Yaskawa INFORM job: OVERLAP2.JBI

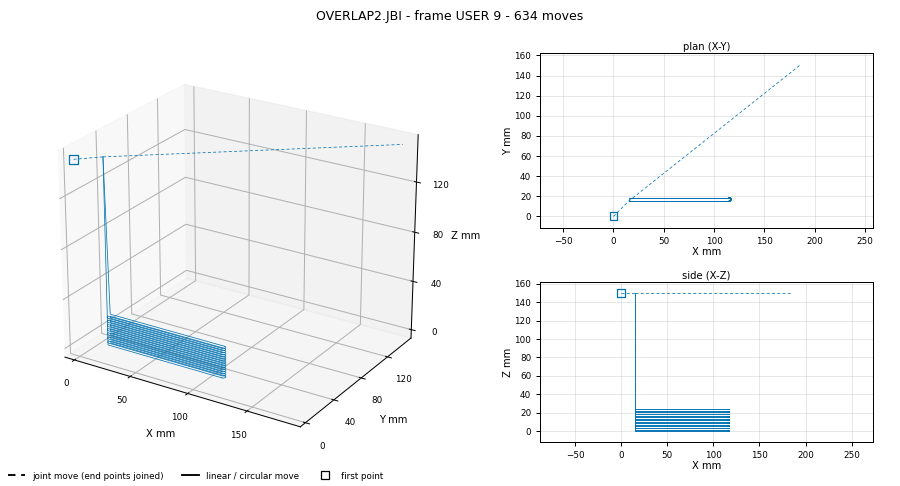
[picture p0: tool path of OVERLAP2.JBI in frame USER 9, 634 of 649 moves have a stored position in this frame; points joined in program order, loops and branches not executed]
/JOB
//NAME OVERLAP1
//POS
///NPOS 649,0,0,0,0,0
///USER 9
///TOOL 1
///POSTYPE USER
///RECTAN
///RCONF 1,0,0,0,0,0,0,0,0,0,0,0,0,0,0,0,0,0,0,0,0,0,0,0
C00000=0.000,0.000,150.000,0.0000,0.0000,-170.0000
C00001=15.000,15.000,150.000,0.0000,0.0000,-170.0000
C00002=15.000,15.000,0.000,0.0000,0.0000,-170.0000
C00003=20.000,15.000,0.000,0.0000,0.0000,-170.0000
C00004=25.000,15.000,0.000,0.0000,0.0000,-170.0000
C00005=30.000,15.000,0.000,0.0000,0.0000,-170.0000
C00006=35.000,15.000,0.000,0.0000,0.0000,-170.0000
C00007=40.000,15.000,0.000,0.0000,0.0000,-170.0000
C00008=45.000,15.000,0.000,0.0000,0.0000,-170.0000
C00009=50.000,15.000,0.000,0.0000,0.0000,-170.0000
C00010=55.000,15.000,0.000,0.0000,0.0000,-170.0000
C00011=60.000,15.000,0.000,0.0000,0.0000,-170.0000
C00012=65.000,15.000,0.000,0.0000,0.0000,-170.0000
C00013=70.000,15.000,0.000,0.0000,0.0000,-170.0000
C00014=75.000,15.000,0.000,0.0000,0.0000,-170.0000
C00015=80.000,15.000,0.000,0.0000,0.0000,-170.0000
C00016=85.000,15.000,0.000,0.0000,0.0000,-170.0000
C00017=90.000,15.000,0.000,0.0000,0.0000,-170.0000
C00018=95.000,15.000,0.000,0.0000,0.0000,-170.0000
C00019=100.000,15.000,0.000,0.0000,0.0000,-170.0000
C00020=105.000,15.000,0.000,0.0000,0.0000,-170.0000
C00021=110.000,15.000,0.000,0.0000,0.0000,-170.0000
C00022=115.000,15.000,0.000,0.0000,0.0000,-170.0000
C00023=116.875,16.875,0.000,0.0000,0.0000,-170.0000
C00024=115.000,18.750,0.000,0.0000,0.0000,-170.0000
C00025=110.000,18.750,0.000,0.0000,0.0000,-170.0000
C00026=105.000,18.750,0.000,0.0000,0.0000,-170.0000
C00027=100.000,18.750,0.000,0.0000,0.0000,-170.0000
C00028=95.000,18.750,0.000,0.0000,0.0000,-170.0000
C00029=90.000,18.750,0.000,0.0000,0.0000,-170.0000
C00030=85.000,18.750,0.000,0.0000,0.0000,-170.0000
C00031=80.000,18.750,0.000,0.0000,0.0000,-170.0000
C00032=75.000,18.750,0.000,0.0000,0.0000,-170.0000
C00033=70.000,18.750,0.000,0.0000,0.0000,-170.0000
C00034=65.000,18.750,0.000,0.0000,0.0000,-170.0000
C00035=60.000,18.750,0.000,0.0000,0.0000,-170.0000
C00036=55.000,18.750,0.000,0.0000,0.0000,-170.0000
C00037=50.000,18.750,0.000,0.0000,0.0000,-170.0000
C00038=45.000,18.750,0.000,0.0000,0.0000,-170.0000
C00039=40.000,18.750,0.000,0.0000,0.0000,-170.0000
C00040=35.000,18.750,0.000,0.0000,0.0000,-170.0000
C00041=30.000,18.750,0.000,0.0000,0.0000,-170.0000
C00042=25.000,18.750,0.000,0.0000,0.0000,-170.0000
C00043=20.000,18.750,0.000,0.0000,0.0000,-170.0000
C00044=15.000,18.750,0.000,0.0000,0.0000,-170.0000
C00045=15.000,18.750,1.700,0.0000,0.0000,-170.0000
C00046=20.000,18.750,1.700,0.0000,0.0000,-170.0000
C00047=25.000,18.750,1.700,0.0000,0.0000,-170.0000
C00048=30.000,18.750,1.700,0.0000,0.0000,-170.0000
C00049=35.000,18.750,1.700,0.0000,0.0000,-170.0000
C00050=40.000,18.750,1.700,0.0000,0.0000,-170.0000
C00051=45.000,18.750,1.700,0.0000,0.0000,-170.0000
C00052=50.000,18.750,1.700,0.0000,0.0000,-170.0000
C00053=55.000,18.750,1.700,0.0000,0.0000,-170.0000
C00054=60.000,18.750,1.700,0.0000,0.0000,-170.0000
C00055=65.000,18.750,1.700,0.0000,0.0000,-170.0000
C00056=70.000,18.750,1.700,0.0000,0.0000,-170.0000
C00057=75.000,18.750,1.700,0.0000,0.0000,-170.0000
C00058=80.000,18.750,1.700,0.0000,0.0000,-170.0000
C00059=85.000,18.750,1.700,0.0000,0.0000,-170.0000
C00060=90.000,18.750,1.700,0.0000,0.0000,-170.0000
C00061=95.000,18.750,1.700,0.0000,0.0000,-170.0000
C00062=100.000,18.750,1.700,0.0000,0.0000,-170.0000
C00063=105.000,18.750,1.700,0.0000,0.0000,-170.0000
C00064=110.000,18.750,1.700,0.0000,0.0000,-170.0000
C00065=115.000,18.750,1.700,0.0000,0.0000,-170.0000
C00066=116.875,16.875,1.700,0.0000,0.0000,-170.0000
C00067=115.000,15.000,1.700,0.0000,0.0000,-170.0000
C00068=110.000,15.000,1.700,0.0000,0.0000,-170.0000
C00069=105.000,15.000,1.700,0.0000,0.0000,-170.0000
C00070=100.000,15.000,1.700,0.0000,0.0000,-170.0000
C00071=95.000,15.000,1.700,0.0000,0.0000,-170.0000
C00072=90.000,15.000,1.700,0.0000,0.0000,-170.0000
C00073=85.000,15.000,1.700,0.0000,0.0000,-170.0000
C00074=80.000,15.000,1.700,0.0000,0.0000,-170.0000
C00075=75.000,15.000,1.700,0.0000,0.0000,-170.0000
C00076=70.000,15.000,1.700,0.0000,0.0000,-170.0000
C00077=65.000,15.000,1.700,0.0000,0.0000,-170.0000
C00078=60.000,15.000,1.700,0.0000,0.0000,-170.0000
C00079=55.000,15.000,1.700,0.0000,0.0000,-170.0000
C00080=50.000,15.000,1.700,0.0000,0.0000,-170.0000
C00081=45.000,15.000,1.700,0.0000,0.0000,-170.0000
C00082=40.000,15.000,1.700,0.0000,0.0000,-170.0000
C00083=35.000,15.000,1.700,0.0000,0.0000,-170.0000
C00084=30.000,15.000,1.700,0.0000,0.0000,-170.0000
C00085=25.000,15.000,1.700,0.0000,0.0000,-170.0000
C00086=20.000,15.000,1.700,0.0000,0.0000,-170.0000
C00087=15.000,15.000,1.700,0.0000,0.0000,-170.0000
C00088=15.000,15.000,3.400,0.0000,0.0000,-170.0000
C00089=20.000,15.000,3.400,0.0000,0.0000,-170.0000
C00090=25.000,15.000,3.400,0.0000,0.0000,-170.0000
C00091=30.000,15.000,3.400,0.0000,0.0000,-170.0000
C00092=35.000,15.000,3.400,0.0000,0.0000,-170.0000
C00093=40.000,15.000,3.400,0.0000,0.0000,-170.0000
C00094=45.000,15.000,3.400,0.0000,0.0000,-170.0000
C00095=50.000,15.000,3.400,0.0000,0.0000,-170.0000
C00096=55.000,15.000,3.400,0.0000,0.0000,-170.0000
C00097=60.000,15.000,3.400,0.0000,0.0000,-170.0000
C00098=65.000,15.000,3.400,0.0000,0.0000,-170.0000
C00099=70.000,15.000,3.400,0.0000,0.0000,-170.0000
C00100=75.000,15.000,3.400,0.0000,0.0000,-170.0000
C00101=80.000,15.000,3.400,0.0000,0.0000,-170.0000
C00102=85.000,15.000,3.400,0.0000,0.0000,-170.0000
C00103=90.000,15.000,3.400,0.0000,0.0000,-170.0000
C00104=95.000,15.000,3.400,0.0000,0.0000,-170.0000
C00105=100.000,15.000,3.400,0.0000,0.0000,-170.0000
C00106=105.000,15.000,3.400,0.0000,0.0000,-170.0000
C00107=110.000,15.000,3.400,0.0000,0.0000,-170.0000
C00108=115.000,15.000,3.400,0.0000,0.0000,-170.0000
C00109=116.875,16.875,3.400,0.0000,0.0000,-170.0000
C00110=115.000,18.750,3.400,0.0000,0.0000,-170.0000
C00111=110.000,18.750,3.400,0.0000,0.0000,-170.0000
C00112=105.000,18.750,3.400,0.0000,0.0000,-170.0000
C00113=100.000,18.750,3.400,0.0000,0.0000,-170.0000
C00114=95.000,18.750,3.400,0.0000,0.0000,-170.0000
C00115=90.000,18.750,3.400,0.0000,0.0000,-170.0000
C00116=85.000,18.750,3.400,0.0000,0.0000,-170.0000
C00117=80.000,18.750,3.400,0.0000,0.0000,-170.0000
C00118=75.000,18.750,3.400,0.0000,0.0000,-170.0000
C00119=70.000,18.750,3.400,0.0000,0.0000,-170.0000
C00120=65.000,18.750,3.400,0.0000,0.0000,-170.0000
C00121=60.000,18.750,3.400,0.0000,0.0000,-170.0000
C00122=55.000,18.750,3.400,0.0000,0.0000,-170.0000
C00123=50.000,18.750,3.400,0.0000,0.0000,-170.0000
C00124=45.000,18.750,3.400,0.0000,0.0000,-170.0000
C00125=40.000,18.750,3.400,0.0000,0.0000,-170.0000
C00126=35.000,18.750,3.400,0.0000,0.0000,-170.0000
C00127=30.000,18.750,3.400,0.0000,0.0000,-170.0000
C00128=25.000,18.750,3.400,0.0000,0.0000,-170.0000
C00129=20.000,18.750,3.400,0.0000,0.0000,-170.0000
C00130=15.000,18.750,3.400,0.0000,0.0000,-170.0000
C00131=15.000,18.750,5.100,0.0000,0.0000,-170.0000
C00132=20.000,18.750,5.100,0.0000,0.0000,-170.0000
C00133=25.000,18.750,5.100,0.0000,0.0000,-170.0000
C00134=30.000,18.750,5.100,0.0000,0.0000,-170.0000
C00135=35.000,18.750,5.100,0.0000,0.0000,-170.0000
C00136=40.000,18.750,5.100,0.0000,0.0000,-170.0000
C00137=45.000,18.750,5.100,0.0000,0.0000,-170.0000
C00138=50.000,18.750,5.100,0.0000,0.0000,-170.0000
C00139=55.000,18.750,5.100,0.0000,0.0000,-170.0000
C00140=60.000,18.750,5.100,0.0000,0.0000,-170.0000
C00141=65.000,18.750,5.100,0.0000,0.0000,-170.0000
C00142=70.000,18.750,5.100,0.0000,0.0000,-170.0000
C00143=75.000,18.750,5.100,0.0000,0.0000,-170.0000
C00144=80.000,18.750,5.100,0.0000,0.0000,-170.0000
C00145=85.000,18.750,5.100,0.0000,0.0000,-170.0000
C00146=90.000,18.750,5.100,0.0000,0.0000,-170.0000
C00147=95.000,18.750,5.100,0.0000,0.0000,-170.0000
C00148=100.000,18.750,5.100,0.0000,0.0000,-170.0000
C00149=105.000,18.750,5.100,0.0000,0.0000,-170.0000
C00150=110.000,18.750,5.100,0.0000,0.0000,-170.0000
C00151=115.000,18.750,5.100,0.0000,0.0000,-170.0000
C00152=116.875,16.875,5.100,0.0000,0.0000,-170.0000
C00153=115.000,15.000,5.100,0.0000,0.0000,-170.0000
C00154=110.000,15.000,5.100,0.0000,0.0000,-170.0000
C00155=105.000,15.000,5.100,0.0000,0.0000,-170.0000
C00156=100.000,15.000,5.100,0.0000,0.0000,-170.0000
C00157=95.000,15.000,5.100,0.0000,0.0000,-170.0000
C00158=90.000,15.000,5.100,0.0000,0.0000,-170.0000
C00159=85.000,15.000,5.100,0.0000,0.0000,-170.0000
C00160=80.000,15.000,5.100,0.0000,0.0000,-170.0000
C00161=75.000,15.000,5.100,0.0000,0.0000,-170.0000
C00162=70.000,15.000,5.100,0.0000,0.0000,-170.0000
C00163=65.000,15.000,5.100,0.0000,0.0000,-170.0000
C00164=60.000,15.000,5.100,0.0000,0.0000,-170.0000
C00165=55.000,15.000,5.100,0.0000,0.0000,-170.0000
C00166=50.000,15.000,5.100,0.0000,0.0000,-170.0000
C00167=45.000,15.000,5.100,0.0000,0.0000,-170.0000
C00168=40.000,15.000,5.100,0.0000,0.0000,-170.0000
C00169=35.000,15.000,5.100,0.0000,0.0000,-170.0000
C00170=30.000,15.000,5.100,0.0000,0.0000,-170.0000
C00171=25.000,15.000,5.100,0.0000,0.0000,-170.0000
C00172=20.000,15.000,5.100,0.0000,0.0000,-170.0000
C00173=15.000,15.000,5.100,0.0000,0.0000,-170.0000
C00174=15.000,15.000,6.800,0.0000,0.0000,-170.0000
C00175=20.000,15.000,6.800,0.0000,0.0000,-170.0000
C00176=25.000,15.000,6.800,0.0000,0.0000,-170.0000
C00177=30.000,15.000,6.800,0.0000,0.0000,-170.0000
C00178=35.000,15.000,6.800,0.0000,0.0000,-170.0000
C00179=40.000,15.000,6.800,0.0000,0.0000,-170.0000
C00180=45.000,15.000,6.800,0.0000,0.0000,-170.0000
C00181=50.000,15.000,6.800,0.0000,0.0000,-170.0000
C00182=55.000,15.000,6.800,0.0000,0.0000,-170.0000
C00183=60.000,15.000,6.800,0.0000,0.0000,-170.0000
C00184=65.000,15.000,6.800,0.0000,0.0000,-170.0000
C00185=70.000,15.000,6.800,0.0000,0.0000,-170.0000
C00186=75.000,15.000,6.800,0.0000,0.0000,-170.0000
C00187=80.000,15.000,6.800,0.0000,0.0000,-170.0000
C00188=85.000,15.000,6.800,0.0000,0.0000,-170.0000
C00189=90.000,15.000,6.800,0.0000,0.0000,-170.0000
C00190=95.000,15.000,6.800,0.0000,0.0000,-170.0000
C00191=100.000,15.000,6.800,0.0000,0.0000,-170.0000
C00192=105.000,15.000,6.800,0.0000,0.0000,-170.0000
C00193=110.000,15.000,6.800,0.0000,0.0000,-170.0000
C00194=115.000,15.000,6.800,0.0000,0.0000,-170.0000
C00195=116.875,16.875,6.800,0.0000,0.0000,-170.0000
C00196=115.000,18.750,6.800,0.0000,0.0000,-170.0000
C00197=110.000,18.750,6.800,0.0000,0.0000,-170.0000
C00198=105.000,18.750,6.800,0.0000,0.0000,-170.0000
C00199=100.000,18.750,6.800,0.0000,0.0000,-170.0000
C00200=95.000,18.750,6.800,0.0000,0.0000,-170.0000
C00201=90.000,18.750,6.800,0.0000,0.0000,-170.0000
C00202=85.000,18.750,6.800,0.0000,0.0000,-170.0000
C00203=80.000,18.750,6.800,0.0000,0.0000,-170.0000
C00204=75.000,18.750,6.800,0.0000,0.0000,-170.0000
C00205=70.000,18.750,6.800,0.0000,0.0000,-170.0000
C00206=65.000,18.750,6.800,0.0000,0.0000,-170.0000
C00207=60.000,18.750,6.800,0.0000,0.0000,-170.0000
C00208=55.000,18.750,6.800,0.0000,0.0000,-170.0000
C00209=50.000,18.750,6.800,0.0000,0.0000,-170.0000
C00210=45.000,18.750,6.800,0.0000,0.0000,-170.0000
C00211=40.000,18.750,6.800,0.0000,0.0000,-170.0000
C00212=35.000,18.750,6.800,0.0000,0.0000,-170.0000
C00213=30.000,18.750,6.800,0.0000,0.0000,-170.0000
C00214=25.000,18.750,6.800,0.0000,0.0000,-170.0000
C00215=20.000,18.750,6.800,0.0000,0.0000,-170.0000
C00216=15.000,18.750,6.800,0.0000,0.0000,-170.0000
C00217=15.000,18.750,8.500,0.0000,0.0000,-170.0000
C00218=20.000,18.750,8.500,0.0000,0.0000,-170.0000
C00219=25.000,18.750,8.500,0.0000,0.0000,-170.0000
C00220=30.000,18.750,8.500,0.0000,0.0000,-170.0000
C00221=35.000,18.750,8.500,0.0000,0.0000,-170.0000
C00222=40.000,18.750,8.500,0.0000,0.0000,-170.0000
C00223=45.000,18.750,8.500,0.0000,0.0000,-170.0000
C00224=50.000,18.750,8.500,0.0000,0.0000,-170.0000
C00225=55.000,18.750,8.500,0.0000,0.0000,-170.0000
C00226=60.000,18.750,8.500,0.0000,0.0000,-170.0000
C00227=65.000,18.750,8.500,0.0000,0.0000,-170.0000
C00228=70.000,18.750,8.500,0.0000,0.0000,-170.0000
C00229=75.000,18.750,8.500,0.0000,0.0000,-170.0000
C00230=80.000,18.750,8.500,0.0000,0.0000,-170.0000
C00231=85.000,18.750,8.500,0.0000,0.0000,-170.0000
C00232=90.000,18.750,8.500,0.0000,0.0000,-170.0000
C00233=95.000,18.750,8.500,0.0000,0.0000,-170.0000
C00234=100.000,18.750,8.500,0.0000,0.0000,-170.0000
C00235=105.000,18.750,8.500,0.0000,0.0000,-170.0000
C00236=110.000,18.750,8.500,0.0000,0.0000,-170.0000
C00237=115.000,18.750,8.500,0.0000,0.0000,-170.0000
C00238=116.875,16.875,8.500,0.0000,0.0000,-170.0000
C00239=115.000,15.000,8.500,0.0000,0.0000,-170.0000
C00240=110.000,15.000,8.500,0.0000,0.0000,-170.0000
C00241=105.000,15.000,8.500,0.0000,0.0000,-170.0000
C00242=100.000,15.000,8.500,0.0000,0.0000,-170.0000
C00243=95.000,15.000,8.500,0.0000,0.0000,-170.0000
C00244=90.000,15.000,8.500,0.0000,0.0000,-170.0000
C00245=85.000,15.000,8.500,0.0000,0.0000,-170.0000
C00246=80.000,15.000,8.500,0.0000,0.0000,-170.0000
C00247=75.000,15.000,8.500,0.0000,0.0000,-170.0000
C00248=70.000,15.000,8.500,0.0000,0.0000,-170.0000
C00249=65.000,15.000,8.500,0.0000,0.0000,-170.0000
C00250=60.000,15.000,8.500,0.0000,0.0000,-170.0000
C00251=55.000,15.000,8.500,0.0000,0.0000,-170.0000
C00252=50.000,15.000,8.500,0.0000,0.0000,-170.0000
C00253=45.000,15.000,8.500,0.0000,0.0000,-170.0000
C00254=40.000,15.000,8.500,0.0000,0.0000,-170.0000
C00255=35.000,15.000,8.500,0.0000,0.0000,-170.0000
C00256=30.000,15.000,8.500,0.0000,0.0000,-170.0000
C00257=25.000,15.000,8.500,0.0000,0.0000,-170.0000
C00258=20.000,15.000,8.500,0.0000,0.0000,-170.0000
C00259=15.000,15.000,8.500,0.0000,0.0000,-170.0000
C00260=15.000,15.000,10.200,0.0000,0.0000,-170.0000
C00261=20.000,15.000,10.200,0.0000,0.0000,-170.0000
C00262=25.000,15.000,10.200,0.0000,0.0000,-170.0000
C00263=30.000,15.000,10.200,0.0000,0.0000,-170.0000
C00264=35.000,15.000,10.200,0.0000,0.0000,-170.0000
C00265=40.000,15.000,10.200,0.0000,0.0000,-170.0000
C00266=45.000,15.000,10.200,0.0000,0.0000,-170.0000
C00267=50.000,15.000,10.200,0.0000,0.0000,-170.0000
C00268=55.000,15.000,10.200,0.0000,0.0000,-170.0000
C00269=60.000,15.000,10.200,0.0000,0.0000,-170.0000
C00270=65.000,15.000,10.200,0.0000,0.0000,-170.0000
C00271=70.000,15.000,10.200,0.0000,0.0000,-170.0000
C00272=75.000,15.000,10.200,0.0000,0.0000,-170.0000
C00273=80.000,15.000,10.200,0.0000,0.0000,-170.0000
C00274=85.000,15.000,10.200,0.0000,0.0000,-170.0000
C00275=90.000,15.000,10.200,0.0000,0.0000,-170.0000
C00276=95.000,15.000,10.200,0.0000,0.0000,-170.0000
C00277=100.000,15.000,10.200,0.0000,0.0000,-170.0000
C00278=105.000,15.000,10.200,0.0000,0.0000,-170.0000
C00279=110.000,15.000,10.200,0.0000,0.0000,-170.0000
C00280=115.000,15.000,10.200,0.0000,0.0000,-170.0000
C00281=116.875,16.875,10.200,0.0000,0.0000,-170.0000
C00282=115.000,18.750,10.200,0.0000,0.0000,-170.0000
C00283=110.000,18.750,10.200,0.0000,0.0000,-170.0000
C00284=105.000,18.750,10.200,0.0000,0.0000,-170.0000
C00285=100.000,18.750,10.200,0.0000,0.0000,-170.0000
C00286=95.000,18.750,10.200,0.0000,0.0000,-170.0000
C00287=90.000,18.750,10.200,0.0000,0.0000,-170.0000
C00288=85.000,18.750,10.200,0.0000,0.0000,-170.0000
C00289=80.000,18.750,10.200,0.0000,0.0000,-170.0000
C00290=75.000,18.750,10.200,0.0000,0.0000,-170.0000
C00291=70.000,18.750,10.200,0.0000,0.0000,-170.0000
C00292=65.000,18.750,10.200,0.0000,0.0000,-170.0000
C00293=60.000,18.750,10.200,0.0000,0.0000,-170.0000
C00294=55.000,18.750,10.200,0.0000,0.0000,-170.0000
C00295=50.000,18.750,10.200,0.0000,0.0000,-170.0000
C00296=45.000,18.750,10.200,0.0000,0.0000,-170.0000
C00297=40.000,18.750,10.200,0.0000,0.0000,-170.0000
C00298=35.000,18.750,10.200,0.0000,0.0000,-170.0000
C00299=30.000,18.750,10.200,0.0000,0.0000,-170.0000
C00300=25.000,18.750,10.200,0.0000,0.0000,-170.0000
C00301=20.000,18.750,10.200,0.0000,0.0000,-170.0000
C00302=15.000,18.750,10.200,0.0000,0.0000,-170.0000
C00303=15.000,18.750,11.900,0.0000,0.0000,-170.0000
C00304=20.000,18.750,11.900,0.0000,0.0000,-170.0000
C00305=25.000,18.750,11.900,0.0000,0.0000,-170.0000
C00306=30.000,18.750,11.900,0.0000,0.0000,-170.0000
C00307=35.000,18.750,11.900,0.0000,0.0000,-170.0000
C00308=40.000,18.750,11.900,0.0000,0.0000,-170.0000
C00309=45.000,18.750,11.900,0.0000,0.0000,-170.0000
C00310=50.000,18.750,11.900,0.0000,0.0000,-170.0000
C00311=55.000,18.750,11.900,0.0000,0.0000,-170.0000
C00312=60.000,18.750,11.900,0.0000,0.0000,-170.0000
C00313=65.000,18.750,11.900,0.0000,0.0000,-170.0000
C00314=70.000,18.750,11.900,0.0000,0.0000,-170.0000
C00315=75.000,18.750,11.900,0.0000,0.0000,-170.0000
C00316=80.000,18.750,11.900,0.0000,0.0000,-170.0000
C00317=85.000,18.750,11.900,0.0000,0.0000,-170.0000
C00318=90.000,18.750,11.900,0.0000,0.0000,-170.0000
C00319=95.000,18.750,11.900,0.0000,0.0000,-170.0000
C00320=100.000,18.750,11.900,0.0000,0.0000,-170.0000
C00321=105.000,18.750,11.900,0.0000,0.0000,-170.0000
C00322=110.000,18.750,11.900,0.0000,0.0000,-170.0000
C00323=115.000,18.750,11.900,0.0000,0.0000,-170.0000
C00324=116.875,16.875,11.900,0.0000,0.0000,-170.0000
C00325=115.000,15.000,11.900,0.0000,0.0000,-170.0000
C00326=110.000,15.000,11.900,0.0000,0.0000,-170.0000
C00327=105.000,15.000,11.900,0.0000,0.0000,-170.0000
C00328=100.000,15.000,11.900,0.0000,0.0000,-170.0000
C00329=95.000,15.000,11.900,0.0000,0.0000,-170.0000
C00330=90.000,15.000,11.900,0.0000,0.0000,-170.0000
C00331=85.000,15.000,11.900,0.0000,0.0000,-170.0000
C00332=80.000,15.000,11.900,0.0000,0.0000,-170.0000
C00333=75.000,15.000,11.900,0.0000,0.0000,-170.0000
C00334=70.000,15.000,11.900,0.0000,0.0000,-170.0000
C00335=65.000,15.000,11.900,0.0000,0.0000,-170.0000
C00336=60.000,15.000,11.900,0.0000,0.0000,-170.0000
C00337=55.000,15.000,11.900,0.0000,0.0000,-170.0000
C00338=50.000,15.000,11.900,0.0000,0.0000,-170.0000
C00339=45.000,15.000,11.900,0.0000,0.0000,-170.0000
C00340=40.000,15.000,11.900,0.0000,0.0000,-170.0000
C00341=35.000,15.000,11.900,0.0000,0.0000,-170.0000
C00342=30.000,15.000,11.900,0.0000,0.0000,-170.0000
C00343=25.000,15.000,11.900,0.0000,0.0000,-170.0000
C00344=20.000,15.000,11.900,0.0000,0.0000,-170.0000
C00345=15.000,15.000,11.900,0.0000,0.0000,-170.0000
C00346=15.000,15.000,13.600,0.0000,0.0000,-170.0000
C00347=20.000,15.000,13.600,0.0000,0.0000,-170.0000
C00348=25.000,15.000,13.600,0.0000,0.0000,-170.0000
C00349=30.000,15.000,13.600,0.0000,0.0000,-170.0000
C00350=35.000,15.000,13.600,0.0000,0.0000,-170.0000
C00351=40.000,15.000,13.600,0.0000,0.0000,-170.0000
C00352=45.000,15.000,13.600,0.0000,0.0000,-170.0000
C00353=50.000,15.000,13.600,0.0000,0.0000,-170.0000
C00354=55.000,15.000,13.600,0.0000,0.0000,-170.0000
C00355=60.000,15.000,13.600,0.0000,0.0000,-170.0000
C00356=65.000,15.000,13.600,0.0000,0.0000,-170.0000
C00357=70.000,15.000,13.600,0.0000,0.0000,-170.0000
C00358=75.000,15.000,13.600,0.0000,0.0000,-170.0000
C00359=80.000,15.000,13.600,0.0000,0.0000,-170.0000
C00360=85.000,15.000,13.600,0.0000,0.0000,-170.0000
C00361=90.000,15.000,13.600,0.0000,0.0000,-170.0000
C00362=95.000,15.000,13.600,0.0000,0.0000,-170.0000
C00363=100.000,15.000,13.600,0.0000,0.0000,-170.0000
C00364=105.000,15.000,13.600,0.0000,0.0000,-170.0000
C00365=110.000,15.000,13.600,0.0000,0.0000,-170.0000
C00366=115.000,15.000,13.600,0.0000,0.0000,-170.0000
C00367=116.875,16.875,13.600,0.0000,0.0000,-170.0000
C00368=115.000,18.750,13.600,0.0000,0.0000,-170.0000
C00369=110.000,18.750,13.600,0.0000,0.0000,-170.0000
C00370=105.000,18.750,13.600,0.0000,0.0000,-170.0000
C00371=100.000,18.750,13.600,0.0000,0.0000,-170.0000
C00372=95.000,18.750,13.600,0.0000,0.0000,-170.0000
C00373=90.000,18.750,13.600,0.0000,0.0000,-170.0000
C00374=85.000,18.750,13.600,0.0000,0.0000,-170.0000
C00375=80.000,18.750,13.600,0.0000,0.0000,-170.0000
C00376=75.000,18.750,13.600,0.0000,0.0000,-170.0000
C00377=70.000,18.750,13.600,0.0000,0.0000,-170.0000
C00378=65.000,18.750,13.600,0.0000,0.0000,-170.0000
C00379=60.000,18.750,13.600,0.0000,0.0000,-170.0000
C00380=55.000,18.750,13.600,0.0000,0.0000,-170.0000
C00381=50.000,18.750,13.600,0.0000,0.0000,-170.0000
C00382=45.000,18.750,13.600,0.0000,0.0000,-170.0000
C00383=40.000,18.750,13.600,0.0000,0.0000,-170.0000
C00384=35.000,18.750,13.600,0.0000,0.0000,-170.0000
C00385=30.000,18.750,13.600,0.0000,0.0000,-170.0000
C00386=25.000,18.750,13.600,0.0000,0.0000,-170.0000
C00387=20.000,18.750,13.600,0.0000,0.0000,-170.0000
C00388=15.000,18.750,13.600,0.0000,0.0000,-170.0000
C00389=15.000,18.750,15.300,0.0000,0.0000,-170.0000
C00390=20.000,18.750,15.300,0.0000,0.0000,-170.0000
C00391=25.000,18.750,15.300,0.0000,0.0000,-170.0000
C00392=30.000,18.750,15.300,0.0000,0.0000,-170.0000
C00393=35.000,18.750,15.300,0.0000,0.0000,-170.0000
C00394=40.000,18.750,15.300,0.0000,0.0000,-170.0000
C00395=45.000,18.750,15.300,0.0000,0.0000,-170.0000
C00396=50.000,18.750,15.300,0.0000,0.0000,-170.0000
C00397=55.000,18.750,15.300,0.0000,0.0000,-170.0000
C00398=60.000,18.750,15.300,0.0000,0.0000,-170.0000
C00399=65.000,18.750,15.300,0.0000,0.0000,-170.0000
C00400=70.000,18.750,15.300,0.0000,0.0000,-170.0000
C00401=75.000,18.750,15.300,0.0000,0.0000,-170.0000
C00402=80.000,18.750,15.300,0.0000,0.0000,-170.0000
C00403=85.000,18.750,15.300,0.0000,0.0000,-170.0000
C00404=90.000,18.750,15.300,0.0000,0.0000,-170.0000
C00405=95.000,18.750,15.300,0.0000,0.0000,-170.0000
C00406=100.000,18.750,15.300,0.0000,0.0000,-170.0000
C00407=105.000,18.750,15.300,0.0000,0.0000,-170.0000
C00408=110.000,18.750,15.300,0.0000,0.0000,-170.0000
C00409=115.000,18.750,15.300,0.0000,0.0000,-170.0000
C00410=116.875,16.875,15.300,0.0000,0.0000,-170.0000
C00411=115.000,15.000,15.300,0.0000,0.0000,-170.0000
C00412=110.000,15.000,15.300,0.0000,0.0000,-170.0000
C00413=105.000,15.000,15.300,0.0000,0.0000,-170.0000
C00414=100.000,15.000,15.300,0.0000,0.0000,-170.0000
C00415=95.000,15.000,15.300,0.0000,0.0000,-170.0000
C00416=90.000,15.000,15.300,0.0000,0.0000,-170.0000
C00417=85.000,15.000,15.300,0.0000,0.0000,-170.0000
C00418=80.000,15.000,15.300,0.0000,0.0000,-170.0000
C00419=75.000,15.000,15.300,0.0000,0.0000,-170.0000
C00420=70.000,15.000,15.300,0.0000,0.0000,-170.0000
C00421=65.000,15.000,15.300,0.0000,0.0000,-170.0000
C00422=60.000,15.000,15.300,0.0000,0.0000,-170.0000
C00423=55.000,15.000,15.300,0.0000,0.0000,-170.0000
C00424=50.000,15.000,15.300,0.0000,0.0000,-170.0000
C00425=45.000,15.000,15.300,0.0000,0.0000,-170.0000
C00426=40.000,15.000,15.300,0.0000,0.0000,-170.0000
C00427=35.000,15.000,15.300,0.0000,0.0000,-170.0000
C00428=30.000,15.000,15.300,0.0000,0.0000,-170.0000
C00429=25.000,15.000,15.300,0.0000,0.0000,-170.0000
C00430=20.000,15.000,15.300,0.0000,0.0000,-170.0000
C00431=15.000,15.000,15.300,0.0000,0.0000,-170.0000
C00432=15.000,15.000,17.000,0.0000,0.0000,-170.0000
C00433=20.000,15.000,17.000,0.0000,0.0000,-170.0000
C00434=25.000,15.000,17.000,0.0000,0.0000,-170.0000
C00435=30.000,15.000,17.000,0.0000,0.0000,-170.0000
C00436=35.000,15.000,17.000,0.0000,0.0000,-170.0000
C00437=40.000,15.000,17.000,0.0000,0.0000,-170.0000
C00438=45.000,15.000,17.000,0.0000,0.0000,-170.0000
C00439=50.000,15.000,17.000,0.0000,0.0000,-170.0000
C00440=55.000,15.000,17.000,0.0000,0.0000,-170.0000
C00441=60.000,15.000,17.000,0.0000,0.0000,-170.0000
C00442=65.000,15.000,17.000,0.0000,0.0000,-170.0000
C00443=70.000,15.000,17.000,0.0000,0.0000,-170.0000
C00444=75.000,15.000,17.000,0.0000,0.0000,-170.0000
C00445=80.000,15.000,17.000,0.0000,0.0000,-170.0000
C00446=85.000,15.000,17.000,0.0000,0.0000,-170.0000
C00447=90.000,15.000,17.000,0.0000,0.0000,-170.0000
C00448=95.000,15.000,17.000,0.0000,0.0000,-170.0000
C00449=100.000,15.000,17.000,0.0000,0.0000,-170.0000
C00450=105.000,15.000,17.000,0.0000,0.0000,-170.0000
C00451=110.000,15.000,17.000,0.0000,0.0000,-170.0000
C00452=115.000,15.000,17.000,0.0000,0.0000,-170.0000
C00453=116.875,16.875,17.000,0.0000,0.0000,-170.0000
C00454=115.000,18.750,17.000,0.0000,0.0000,-170.0000
C00455=110.000,18.750,17.000,0.0000,0.0000,-170.0000
C00456=105.000,18.750,17.000,0.0000,0.0000,-170.0000
C00457=100.000,18.750,17.000,0.0000,0.0000,-170.0000
C00458=95.000,18.750,17.000,0.0000,0.0000,-170.0000
C00459=90.000,18.750,17.000,0.0000,0.0000,-170.0000
C00460=85.000,18.750,17.000,0.0000,0.0000,-170.0000
C00461=80.000,18.750,17.000,0.0000,0.0000,-170.0000
C00462=75.000,18.750,17.000,0.0000,0.0000,-170.0000
C00463=70.000,18.750,17.000,0.0000,0.0000,-170.0000
C00464=65.000,18.750,17.000,0.0000,0.0000,-170.0000
C00465=60.000,18.750,17.000,0.0000,0.0000,-170.0000
C00466=55.000,18.750,17.000,0.0000,0.0000,-170.0000
C00467=50.000,18.750,17.000,0.0000,0.0000,-170.0000
C00468=45.000,18.750,17.000,0.0000,0.0000,-170.0000
C00469=40.000,18.750,17.000,0.0000,0.0000,-170.0000
C00470=35.000,18.750,17.000,0.0000,0.0000,-170.0000
C00471=30.000,18.750,17.000,0.0000,0.0000,-170.0000
C00472=25.000,18.750,17.000,0.0000,0.0000,-170.0000
C00473=20.000,18.750,17.000,0.0000,0.0000,-170.0000
C00474=15.000,18.750,17.000,0.0000,0.0000,-170.0000
C00475=15.000,18.750,18.700,0.0000,0.0000,-170.0000
C00476=20.000,18.750,18.700,0.0000,0.0000,-170.0000
C00477=25.000,18.750,18.700,0.0000,0.0000,-170.0000
C00478=30.000,18.750,18.700,0.0000,0.0000,-170.0000
C00479=35.000,18.750,18.700,0.0000,0.0000,-170.0000
C00480=40.000,18.750,18.700,0.0000,0.0000,-170.0000
C00481=45.000,18.750,18.700,0.0000,0.0000,-170.0000
C00482=50.000,18.750,18.700,0.0000,0.0000,-170.0000
C00483=55.000,18.750,18.700,0.0000,0.0000,-170.0000
C00484=60.000,18.750,18.700,0.0000,0.0000,-170.0000
C00485=65.000,18.750,18.700,0.0000,0.0000,-170.0000
C00486=70.000,18.750,18.700,0.0000,0.0000,-170.0000
C00487=75.000,18.750,18.700,0.0000,0.0000,-170.0000
C00488=80.000,18.750,18.700,0.0000,0.0000,-170.0000
C00489=85.000,18.750,18.700,0.0000,0.0000,-170.0000
C00490=90.000,18.750,18.700,0.0000,0.0000,-170.0000
C00491=95.000,18.750,18.700,0.0000,0.0000,-170.0000
C00492=100.000,18.750,18.700,0.0000,0.0000,-170.0000
C00493=105.000,18.750,18.700,0.0000,0.0000,-170.0000
C00494=110.000,18.750,18.700,0.0000,0.0000,-170.0000
C00495=115.000,18.750,18.700,0.0000,0.0000,-170.0000
C00496=116.875,16.875,18.700,0.0000,0.0000,-170.0000
C00497=115.000,15.000,18.700,0.0000,0.0000,-170.0000
C00498=110.000,15.000,18.700,0.0000,0.0000,-170.0000
C00499=105.000,15.000,18.700,0.0000,0.0000,-170.0000
C00500=100.000,15.000,18.700,0.0000,0.0000,-170.0000
C00501=95.000,15.000,18.700,0.0000,0.0000,-170.0000
C00502=90.000,15.000,18.700,0.0000,0.0000,-170.0000
C00503=85.000,15.000,18.700,0.0000,0.0000,-170.0000
C00504=80.000,15.000,18.700,0.0000,0.0000,-170.0000
C00505=75.000,15.000,18.700,0.0000,0.0000,-170.0000
C00506=70.000,15.000,18.700,0.0000,0.0000,-170.0000
C00507=65.000,15.000,18.700,0.0000,0.0000,-170.0000
C00508=60.000,15.000,18.700,0.0000,0.0000,-170.0000
C00509=55.000,15.000,18.700,0.0000,0.0000,-170.0000
C00510=50.000,15.000,18.700,0.0000,0.0000,-170.0000
C00511=45.000,15.000,18.700,0.0000,0.0000,-170.0000
C00512=40.000,15.000,18.700,0.0000,0.0000,-170.0000
C00513=35.000,15.000,18.700,0.0000,0.0000,-170.0000
C00514=30.000,15.000,18.700,0.0000,0.0000,-170.0000
C00515=25.000,15.000,18.700,0.0000,0.0000,-170.0000
C00516=20.000,15.000,18.700,0.0000,0.0000,-170.0000
C00517=15.000,15.000,18.700,0.0000,0.0000,-170.0000
C00518=15.000,15.000,20.400,0.0000,0.0000,-170.0000
C00519=20.000,15.000,20.400,0.0000,0.0000,-170.0000
C00520=25.000,15.000,20.400,0.0000,0.0000,-170.0000
C00521=30.000,15.000,20.400,0.0000,0.0000,-170.0000
C00522=35.000,15.000,20.400,0.0000,0.0000,-170.0000
C00523=40.000,15.000,20.400,0.0000,0.0000,-170.0000
C00524=45.000,15.000,20.400,0.0000,0.0000,-170.0000
C00525=50.000,15.000,20.400,0.0000,0.0000,-170.0000
C00526=55.000,15.000,20.400,0.0000,0.0000,-170.0000
C00527=60.000,15.000,20.400,0.0000,0.0000,-170.0000
C00528=65.000,15.000,20.400,0.0000,0.0000,-170.0000
C00529=70.000,15.000,20.400,0.0000,0.0000,-170.0000
C00530=75.000,15.000,20.400,0.0000,0.0000,-170.0000
C00531=80.000,15.000,20.400,0.0000,0.0000,-170.0000
C00532=85.000,15.000,20.400,0.0000,0.0000,-170.0000
C00533=90.000,15.000,20.400,0.0000,0.0000,-170.0000
C00534=95.000,15.000,20.400,0.0000,0.0000,-170.0000
C00535=100.000,15.000,20.400,0.0000,0.0000,-170.0000
C00536=105.000,15.000,20.400,0.0000,0.0000,-170.0000
C00537=110.000,15.000,20.400,0.0000,0.0000,-170.0000
C00538=115.000,15.000,20.400,0.0000,0.0000,-170.0000
C00539=116.875,16.875,20.400,0.0000,0.0000,-170.0000
C00540=115.000,18.750,20.400,0.0000,0.0000,-170.0000
C00541=110.000,18.750,20.400,0.0000,0.0000,-170.0000
C00542=105.000,18.750,20.400,0.0000,0.0000,-170.0000
C00543=100.000,18.750,20.400,0.0000,0.0000,-170.0000
C00544=95.000,18.750,20.400,0.0000,0.0000,-170.0000
C00545=90.000,18.750,20.400,0.0000,0.0000,-170.0000
C00546=85.000,18.750,20.400,0.0000,0.0000,-170.0000
C00547=80.000,18.750,20.400,0.0000,0.0000,-170.0000
C00548=75.000,18.750,20.400,0.0000,0.0000,-170.0000
C00549=70.000,18.750,20.400,0.0000,0.0000,-170.0000
C00550=65.000,18.750,20.400,0.0000,0.0000,-170.0000
C00551=60.000,18.750,20.400,0.0000,0.0000,-170.0000
C00552=55.000,18.750,20.400,0.0000,0.0000,-170.0000
C00553=50.000,18.750,20.400,0.0000,0.0000,-170.0000
C00554=45.000,18.750,20.400,0.0000,0.0000,-170.0000
C00555=40.000,18.750,20.400,0.0000,0.0000,-170.0000
C00556=35.000,18.750,20.400,0.0000,0.0000,-170.0000
C00557=30.000,18.750,20.400,0.0000,0.0000,-170.0000
C00558=25.000,18.750,20.400,0.0000,0.0000,-170.0000
C00559=20.000,18.750,20.400,0.0000,0.0000,-170.0000
C00560=15.000,18.750,20.400,0.0000,0.0000,-170.0000
C00561=15.000,18.750,22.100,0.0000,0.0000,-170.0000
C00562=20.000,18.750,22.100,0.0000,0.0000,-170.0000
C00563=25.000,18.750,22.100,0.0000,0.0000,-170.0000
C00564=30.000,18.750,22.100,0.0000,0.0000,-170.0000
C00565=35.000,18.750,22.100,0.0000,0.0000,-170.0000
C00566=40.000,18.750,22.100,0.0000,0.0000,-170.0000
C00567=45.000,18.750,22.100,0.0000,0.0000,-170.0000
C00568=50.000,18.750,22.100,0.0000,0.0000,-170.0000
C00569=55.000,18.750,22.100,0.0000,0.0000,-170.0000
C00570=60.000,18.750,22.100,0.0000,0.0000,-170.0000
C00571=65.000,18.750,22.100,0.0000,0.0000,-170.0000
C00572=70.000,18.750,22.100,0.0000,0.0000,-170.0000
C00573=75.000,18.750,22.100,0.0000,0.0000,-170.0000
C00574=80.000,18.750,22.100,0.0000,0.0000,-170.0000
C00575=85.000,18.750,22.100,0.0000,0.0000,-170.0000
C00576=90.000,18.750,22.100,0.0000,0.0000,-170.0000
C00577=95.000,18.750,22.100,0.0000,0.0000,-170.0000
C00578=100.000,18.750,22.100,0.0000,0.0000,-170.0000
C00579=105.000,18.750,22.100,0.0000,0.0000,-170.0000
C00580=110.000,18.750,22.100,0.0000,0.0000,-170.0000
C00581=115.000,18.750,22.100,0.0000,0.0000,-170.0000
C00582=116.875,16.875,22.100,0.0000,0.0000,-170.0000
C00583=115.000,15.000,22.100,0.0000,0.0000,-170.0000
C00584=110.000,15.000,22.100,0.0000,0.0000,-170.0000
C00585=105.000,15.000,22.100,0.0000,0.0000,-170.0000
C00586=100.000,15.000,22.100,0.0000,0.0000,-170.0000
C00587=95.000,15.000,22.100,0.0000,0.0000,-170.0000
C00588=90.000,15.000,22.100,0.0000,0.0000,-170.0000
C00589=85.000,15.000,22.100,0.0000,0.0000,-170.0000
C00590=80.000,15.000,22.100,0.0000,0.0000,-170.0000
C00591=75.000,15.000,22.100,0.0000,0.0000,-170.0000
C00592=70.000,15.000,22.100,0.0000,0.0000,-170.0000
C00593=65.000,15.000,22.100,0.0000,0.0000,-170.0000
C00594=60.000,15.000,22.100,0.0000,0.0000,-170.0000
C00595=55.000,15.000,22.100,0.0000,0.0000,-170.0000
C00596=50.000,15.000,22.100,0.0000,0.0000,-170.0000
C00597=45.000,15.000,22.100,0.0000,0.0000,-170.0000
C00598=40.000,15.000,22.100,0.0000,0.0000,-170.0000
C00599=35.000,15.000,22.100,0.0000,0.0000,-170.0000
C00600=30.000,15.000,22.100,0.0000,0.0000,-170.0000
C00601=25.000,15.000,22.100,0.0000,0.0000,-170.0000
C00602=20.000,15.000,22.100,0.0000,0.0000,-170.0000
C00603=15.000,15.000,22.100,0.0000,0.0000,-170.0000
C00604=15.000,15.000,23.800,0.0000,0.0000,-170.0000
C00605=20.000,15.000,23.800,0.0000,0.0000,-170.0000
C00606=25.000,15.000,23.800,0.0000,0.0000,-170.0000
C00607=30.000,15.000,23.800,0.0000,0.0000,-170.0000
C00608=35.000,15.000,23.800,0.0000,0.0000,-170.0000
C00609=40.000,15.000,23.800,0.0000,0.0000,-170.0000
C00610=45.000,15.000,23.800,0.0000,0.0000,-170.0000
C00611=50.000,15.000,23.800,0.0000,0.0000,-170.0000
C00612=55.000,15.000,23.800,0.0000,0.0000,-170.0000
C00613=60.000,15.000,23.800,0.0000,0.0000,-170.0000
C00614=65.000,15.000,23.800,0.0000,0.0000,-170.0000
C00615=70.000,15.000,23.800,0.0000,0.0000,-170.0000
C00616=75.000,15.000,23.800,0.0000,0.0000,-170.0000
C00617=80.000,15.000,23.800,0.0000,0.0000,-170.0000
C00618=85.000,15.000,23.800,0.0000,0.0000,-170.0000
C00619=90.000,15.000,23.800,0.0000,0.0000,-170.0000
C00620=95.000,15.000,23.800,0.0000,0.0000,-170.0000
C00621=100.000,15.000,23.800,0.0000,0.0000,-170.0000
C00622=105.000,15.000,23.800,0.0000,0.0000,-170.0000
C00623=110.000,15.000,23.800,0.0000,0.0000,-170.0000
C00624=115.000,15.000,23.800,0.0000,0.0000,-170.0000
C00625=116.875,16.875,23.800,0.0000,0.0000,-170.0000
C00626=115.000,18.750,23.800,0.0000,0.0000,-170.0000
C00627=110.000,18.750,23.800,0.0000,0.0000,-170.0000
C00628=105.000,18.750,23.800,0.0000,0.0000,-170.0000
C00629=100.000,18.750,23.800,0.0000,0.0000,-170.0000
C00630=95.000,18.750,23.800,0.0000,0.0000,-170.0000
C00631=90.000,18.750,23.800,0.0000,0.0000,-170.0000
C00632=85.000,18.750,23.800,0.0000,0.0000,-170.0000
C00633=80.000,18.750,23.800,0.0000,0.0000,-170.0000
C00634=75.000,18.750,23.800,0.0000,0.0000,-170.0000
C00635=70.000,18.750,23.800,0.0000,0.0000,-170.0000
C00636=65.000,18.750,23.800,0.0000,0.0000,-170.0000
C00637=60.000,18.750,23.800,0.0000,0.0000,-170.0000
C00638=55.000,18.750,23.800,0.0000,0.0000,-170.0000
C00639=50.000,18.750,23.800,0.0000,0.0000,-170.0000
C00640=45.000,18.750,23.800,0.0000,0.0000,-170.0000
C00641=40.000,18.750,23.800,0.0000,0.0000,-170.0000
C00642=35.000,18.750,23.800,0.0000,0.0000,-170.0000
C00643=30.000,18.750,23.800,0.0000,0.0000,-170.0000
C00644=25.000,18.750,23.800,0.0000,0.0000,-170.0000
C00645=20.000,18.750,23.800,0.0000,0.0000,-170.0000
C00646=15.000,18.750,23.800,0.0000,0.0000,-170.0000
C00647=15.000,15.000,150.000,0.0000,0.0000,-170.0000
C00648=185.000,150.000,150.000,0.0000,0.0000,-170.0000
//INST
///DATE 2026/11/06 13:28
///ATTR SC,RW,RJ
////FRAME USER 9
///GROUP1 RB1
NOP
MOVJ C00000 VJ=0.78
MOVJ C00001 VJ=0.78
MOVL C00002 V=11.0 PL=0
*LAG1
MACRO1 MJ#(0) ARGF1
ARCON
MOVL C00003 V=7.0 PL=0
MOVL C00004 V=7.0 PL=0
MOVL C00005 V=7.0 PL=0
MOVL C00006 V=7.0 PL=0
MOVL C00007 V=7.0 PL=0
MOVL C00008 V=7.0 PL=0
MOVL C00009 V=7.0 PL=0
MOVL C00010 V=7.0 PL=0
MOVL C00011 V=7.0 PL=0
MOVL C00012 V=7.0 PL=0
MOVL C00013 V=7.0 PL=0
MOVL C00014 V=7.0 PL=0
MOVL C00015 V=7.0 PL=0
MOVL C00016 V=7.0 PL=0
MOVL C00017 V=7.0 PL=0
MOVL C00018 V=7.0 PL=0
MOVL C00019 V=7.0 PL=0
MOVL C00020 V=7.0 PL=0
MOVL C00021 V=7.0 PL=0
MOVC C00022 V=7.0 ACC=20 DEC=20
MOVC C00023 V=7.0 ACC=20 DEC=20
MOVC C00024 V=7.0 ACC=20 DEC=20
MOVL C00025 V=7.0 PL=0
MOVL C00026 V=7.0 PL=0
MOVL C00027 V=7.0 PL=0
MOVL C00028 V=7.0 PL=0
MOVL C00029 V=7.0 PL=0
MOVL C00030 V=7.0 PL=0
MOVL C00031 V=7.0 PL=0
MOVL C00032 V=7.0 PL=0
MOVL C00033 V=7.0 PL=0
MOVL C00034 V=7.0 PL=0
MOVL C00035 V=7.0 PL=0
MOVL C00036 V=7.0 PL=0
MOVL C00037 V=7.0 PL=0
MOVL C00038 V=7.0 PL=0
MOVL C00039 V=7.0 PL=0
MOVL C00040 V=7.0 PL=0
MOVL C00041 V=7.0 PL=0
MOVL C00042 V=7.0 PL=0
MOVL C00043 V=7.0 PL=0
MOVL C00044 V=7.0 PL=0
ARCOF
TIMER T=30.00
*LAG2
MOVL C00045 V=11.0 PL=0
MACRO1 MJ#(0) ARGF2
ARCON
MOVL C00046 V=7.0 PL=0
MOVL C00047 V=7.0 PL=0
MOVL C00048 V=7.0 PL=0
MOVL C00049 V=7.0 PL=0
MOVL C00050 V=7.0 PL=0
MOVL C00051 V=7.0 PL=0
MOVL C00052 V=7.0 PL=0
MOVL C00053 V=7.0 PL=0
MOVL C00054 V=7.0 PL=0
MOVL C00055 V=7.0 PL=0
MOVL C00056 V=7.0 PL=0
MOVL C00057 V=7.0 PL=0
MOVL C00058 V=7.0 PL=0
MOVL C00059 V=7.0 PL=0
MOVL C00060 V=7.0 PL=0
MOVL C00061 V=7.0 PL=0
MOVL C00062 V=7.0 PL=0
MOVL C00063 V=7.0 PL=0
MOVL C00064 V=7.0 PL=0
MOVC C00065 V=7.0 ACC=20 DEC=20
MOVC C00066 V=7.0 ACC=20 DEC=20
MOVC C00067 V=7.0 ACC=20 DEC=20
MOVL C00068 V=7.0 PL=0
MOVL C00069 V=7.0 PL=0
MOVL C00070 V=7.0 PL=0
MOVL C00071 V=7.0 PL=0
MOVL C00072 V=7.0 PL=0
MOVL C00073 V=7.0 PL=0
MOVL C00074 V=7.0 PL=0
MOVL C00075 V=7.0 PL=0
MOVL C00076 V=7.0 PL=0
MOVL C00077 V=7.0 PL=0
MOVL C00078 V=7.0 PL=0
MOVL C00079 V=7.0 PL=0
MOVL C00080 V=7.0 PL=0
MOVL C00081 V=7.0 PL=0
MOVL C00082 V=7.0 PL=0
MOVL C00083 V=7.0 PL=0
MOVL C00084 V=7.0 PL=0
MOVL C00085 V=7.0 PL=0
MOVL C00086 V=7.0 PL=0
MOVL C00087 V=7.0 PL=0
ARCOF
TIMER T=30.00
*LAG3
MOVL C00088 V=11.0 PL=0
MACRO1 MJ#(0) ARGF2
ARCON
MOVL C00089 V=7.0 PL=0
MOVL C00090 V=7.0 PL=0
MOVL C00091 V=7.0 PL=0
MOVL C00092 V=7.0 PL=0
MOVL C00093 V=7.0 PL=0
MOVL C00094 V=7.0 PL=0
MOVL C00095 V=7.0 PL=0
MOVL C00096 V=7.0 PL=0
MOVL C00097 V=7.0 PL=0
MOVL C00098 V=7.0 PL=0
MOVL C00099 V=7.0 PL=0
MOVL C00100 V=7.0 PL=0
MOVL C00101 V=7.0 PL=0
MOVL C00102 V=7.0 PL=0
MOVL C00103 V=7.0 PL=0
MOVL C00104 V=7.0 PL=0
MOVL C00105 V=7.0 PL=0
MOVL C00106 V=7.0 PL=0
MOVL C00107 V=7.0 PL=0
MOVC C00108 V=7.0 ACC=20 DEC=20
MOVC C00109 V=7.0 ACC=20 DEC=20
MOVC C00110 V=7.0 ACC=20 DEC=20
MOVL C00111 V=7.0 PL=0
MOVL C00112 V=7.0 PL=0
MOVL C00113 V=7.0 PL=0
MOVL C00114 V=7.0 PL=0
MOVL C00115 V=7.0 PL=0
MOVL C00116 V=7.0 PL=0
MOVL C00117 V=7.0 PL=0
MOVL C00118 V=7.0 PL=0
MOVL C00119 V=7.0 PL=0
MOVL C00120 V=7.0 PL=0
MOVL C00121 V=7.0 PL=0
MOVL C00122 V=7.0 PL=0
MOVL C00123 V=7.0 PL=0
MOVL C00124 V=7.0 PL=0
MOVL C00125 V=7.0 PL=0
MOVL C00126 V=7.0 PL=0
MOVL C00127 V=7.0 PL=0
MOVL C00128 V=7.0 PL=0
MOVL C00129 V=7.0 PL=0
MOVL C00130 V=7.0 PL=0
ARCOF
TIMER T=30.00
*LAG4
MOVL C00131 V=11.0 PL=0
MACRO1 MJ#(0) ARGF2
ARCON
MOVL C00132 V=7.0 PL=0
MOVL C00133 V=7.0 PL=0
MOVL C00134 V=7.0 PL=0
MOVL C00135 V=7.0 PL=0
MOVL C00136 V=7.0 PL=0
MOVL C00137 V=7.0 PL=0
MOVL C00138 V=7.0 PL=0
MOVL C00139 V=7.0 PL=0
MOVL C00140 V=7.0 PL=0
MOVL C00141 V=7.0 PL=0
MOVL C00142 V=7.0 PL=0
MOVL C00143 V=7.0 PL=0
MOVL C00144 V=7.0 PL=0
MOVL C00145 V=7.0 PL=0
MOVL C00146 V=7.0 PL=0
MOVL C00147 V=7.0 PL=0
MOVL C00148 V=7.0 PL=0
MOVL C00149 V=7.0 PL=0
MOVL C00150 V=7.0 PL=0
MOVC C00151 V=7.0 ACC=20 DEC=20
MOVC C00152 V=7.0 ACC=20 DEC=20
MOVC C00153 V=7.0 ACC=20 DEC=20
MOVL C00154 V=7.0 PL=0
MOVL C00155 V=7.0 PL=0
MOVL C00156 V=7.0 PL=0
MOVL C00157 V=7.0 PL=0
MOVL C00158 V=7.0 PL=0
MOVL C00159 V=7.0 PL=0
MOVL C00160 V=7.0 PL=0
MOVL C00161 V=7.0 PL=0
MOVL C00162 V=7.0 PL=0
MOVL C00163 V=7.0 PL=0
MOVL C00164 V=7.0 PL=0
MOVL C00165 V=7.0 PL=0
MOVL C00166 V=7.0 PL=0
MOVL C00167 V=7.0 PL=0
MOVL C00168 V=7.0 PL=0
MOVL C00169 V=7.0 PL=0
MOVL C00170 V=7.0 PL=0
MOVL C00171 V=7.0 PL=0
MOVL C00172 V=7.0 PL=0
MOVL C00173 V=7.0 PL=0
ARCOF
TIMER T=30.00
*LAG5
MOVL C00174 V=11.0 PL=0
MACRO1 MJ#(0) ARGF2
ARCON
MOVL C00175 V=7.0 PL=0
MOVL C00176 V=7.0 PL=0
MOVL C00177 V=7.0 PL=0
MOVL C00178 V=7.0 PL=0
MOVL C00179 V=7.0 PL=0
MOVL C00180 V=7.0 PL=0
MOVL C00181 V=7.0 PL=0
MOVL C00182 V=7.0 PL=0
MOVL C00183 V=7.0 PL=0
MOVL C00184 V=7.0 PL=0
MOVL C00185 V=7.0 PL=0
MOVL C00186 V=7.0 PL=0
MOVL C00187 V=7.0 PL=0
MOVL C00188 V=7.0 PL=0
MOVL C00189 V=7.0 PL=0
MOVL C00190 V=7.0 PL=0
MOVL C00191 V=7.0 PL=0
MOVL C00192 V=7.0 PL=0
MOVL C00193 V=7.0 PL=0
MOVC C00194 V=7.0 ACC=20 DEC=20
MOVC C00195 V=7.0 ACC=20 DEC=20
MOVC C00196 V=7.0 ACC=20 DEC=20
MOVL C00197 V=7.0 PL=0
MOVL C00198 V=7.0 PL=0
MOVL C00199 V=7.0 PL=0
MOVL C00200 V=7.0 PL=0
MOVL C00201 V=7.0 PL=0
MOVL C00202 V=7.0 PL=0
MOVL C00203 V=7.0 PL=0
MOVL C00204 V=7.0 PL=0
MOVL C00205 V=7.0 PL=0
MOVL C00206 V=7.0 PL=0
MOVL C00207 V=7.0 PL=0
MOVL C00208 V=7.0 PL=0
MOVL C00209 V=7.0 PL=0
MOVL C00210 V=7.0 PL=0
MOVL C00211 V=7.0 PL=0
MOVL C00212 V=7.0 PL=0
MOVL C00213 V=7.0 PL=0
MOVL C00214 V=7.0 PL=0
MOVL C00215 V=7.0 PL=0
MOVL C00216 V=7.0 PL=0
ARCOF
TIMER T=30.00
*LAG6
MOVL C00217 V=11.0 PL=0
MACRO1 MJ#(0) ARGF2
ARCON
MOVL C00218 V=7.0 PL=0
MOVL C00219 V=7.0 PL=0
MOVL C00220 V=7.0 PL=0
MOVL C00221 V=7.0 PL=0
MOVL C00222 V=7.0 PL=0
MOVL C00223 V=7.0 PL=0
MOVL C00224 V=7.0 PL=0
MOVL C00225 V=7.0 PL=0
MOVL C00226 V=7.0 PL=0
MOVL C00227 V=7.0 PL=0
MOVL C00228 V=7.0 PL=0
MOVL C00229 V=7.0 PL=0
MOVL C00230 V=7.0 PL=0
MOVL C00231 V=7.0 PL=0
MOVL C00232 V=7.0 PL=0
MOVL C00233 V=7.0 PL=0
MOVL C00234 V=7.0 PL=0
MOVL C00235 V=7.0 PL=0
MOVL C00236 V=7.0 PL=0
MOVC C00237 V=7.0 ACC=20 DEC=20
MOVC C00238 V=7.0 ACC=20 DEC=20
MOVC C00239 V=7.0 ACC=20 DEC=20
MOVL C00240 V=7.0 PL=0
MOVL C00241 V=7.0 PL=0
MOVL C00242 V=7.0 PL=0
MOVL C00243 V=7.0 PL=0
MOVL C00244 V=7.0 PL=0
MOVL C00245 V=7.0 PL=0
MOVL C00246 V=7.0 PL=0
MOVL C00247 V=7.0 PL=0
MOVL C00248 V=7.0 PL=0
MOVL C00249 V=7.0 PL=0
MOVL C00250 V=7.0 PL=0
MOVL C00251 V=7.0 PL=0
MOVL C00252 V=7.0 PL=0
MOVL C00253 V=7.0 PL=0
MOVL C00254 V=7.0 PL=0
MOVL C00255 V=7.0 PL=0
MOVL C00256 V=7.0 PL=0
MOVL C00257 V=7.0 PL=0
MOVL C00258 V=7.0 PL=0
MOVL C00259 V=7.0 PL=0
ARCOF
TIMER T=30.00
*LAG7
MOVL C00260 V=11.0 PL=0
MACRO1 MJ#(0) ARGF2
ARCON
MOVL C00261 V=7.0 PL=0
MOVL C00262 V=7.0 PL=0
MOVL C00263 V=7.0 PL=0
MOVL C00264 V=7.0 PL=0
MOVL C00265 V=7.0 PL=0
MOVL C00266 V=7.0 PL=0
MOVL C00267 V=7.0 PL=0
MOVL C00268 V=7.0 PL=0
MOVL C00269 V=7.0 PL=0
MOVL C00270 V=7.0 PL=0
MOVL C00271 V=7.0 PL=0
MOVL C00272 V=7.0 PL=0
MOVL C00273 V=7.0 PL=0
MOVL C00274 V=7.0 PL=0
MOVL C00275 V=7.0 PL=0
MOVL C00276 V=7.0 PL=0
MOVL C00277 V=7.0 PL=0
MOVL C00278 V=7.0 PL=0
MOVL C00279 V=7.0 PL=0
MOVC C00280 V=7.0 ACC=20 DEC=20
MOVC C00281 V=7.0 ACC=20 DEC=20
MOVC C00282 V=7.0 ACC=20 DEC=20
MOVL C00283 V=7.0 PL=0
MOVL C00284 V=7.0 PL=0
MOVL C00285 V=7.0 PL=0
MOVL C00286 V=7.0 PL=0
MOVL C00287 V=7.0 PL=0
MOVL C00288 V=7.0 PL=0
MOVL C00289 V=7.0 PL=0
MOVL C00290 V=7.0 PL=0
MOVL C00291 V=7.0 PL=0
MOVL C00292 V=7.0 PL=0
MOVL C00293 V=7.0 PL=0
MOVL C00294 V=7.0 PL=0
MOVL C00295 V=7.0 PL=0
MOVL C00296 V=7.0 PL=0
MOVL C00297 V=7.0 PL=0
MOVL C00298 V=7.0 PL=0
MOVL C00299 V=7.0 PL=0
MOVL C00300 V=7.0 PL=0
MOVL C00301 V=7.0 PL=0
MOVL C00302 V=7.0 PL=0
ARCOF
TIMER T=30.00
*LAG8
MOVL C00303 V=11.0 PL=0
MACRO1 MJ#(0) ARGF2
ARCON
MOVL C00304 V=7.0 PL=0
MOVL C00305 V=7.0 PL=0
MOVL C00306 V=7.0 PL=0
MOVL C00307 V=7.0 PL=0
MOVL C00308 V=7.0 PL=0
MOVL C00309 V=7.0 PL=0
MOVL C00310 V=7.0 PL=0
MOVL C00311 V=7.0 PL=0
MOVL C00312 V=7.0 PL=0
MOVL C00313 V=7.0 PL=0
MOVL C00314 V=7.0 PL=0
MOVL C00315 V=7.0 PL=0
MOVL C00316 V=7.0 PL=0
MOVL C00317 V=7.0 PL=0
MOVL C00318 V=7.0 PL=0
MOVL C00319 V=7.0 PL=0
MOVL C00320 V=7.0 PL=0
MOVL C00321 V=7.0 PL=0
MOVL C00322 V=7.0 PL=0
MOVC C00323 V=7.0 ACC=20 DEC=20
MOVC C00324 V=7.0 ACC=20 DEC=20
MOVC C00325 V=7.0 ACC=20 DEC=20
MOVL C00326 V=7.0 PL=0
MOVL C00327 V=7.0 PL=0
MOVL C00328 V=7.0 PL=0
MOVL C00329 V=7.0 PL=0
MOVL C00330 V=7.0 PL=0
MOVL C00331 V=7.0 PL=0
MOVL C00332 V=7.0 PL=0
MOVL C00333 V=7.0 PL=0
MOVL C00334 V=7.0 PL=0
MOVL C00335 V=7.0 PL=0
MOVL C00336 V=7.0 PL=0
MOVL C00337 V=7.0 PL=0
MOVL C00338 V=7.0 PL=0
MOVL C00339 V=7.0 PL=0
MOVL C00340 V=7.0 PL=0
MOVL C00341 V=7.0 PL=0
MOVL C00342 V=7.0 PL=0
MOVL C00343 V=7.0 PL=0
MOVL C00344 V=7.0 PL=0
MOVL C00345 V=7.0 PL=0
ARCOF
TIMER T=30.00
*LAG9
MOVL C00346 V=11.0 PL=0
MACRO1 MJ#(0) ARGF2
ARCON
MOVL C00347 V=7.0 PL=0
MOVL C00348 V=7.0 PL=0
MOVL C00349 V=7.0 PL=0
MOVL C00350 V=7.0 PL=0
MOVL C00351 V=7.0 PL=0
MOVL C00352 V=7.0 PL=0
MOVL C00353 V=7.0 PL=0
MOVL C00354 V=7.0 PL=0
MOVL C00355 V=7.0 PL=0
MOVL C00356 V=7.0 PL=0
MOVL C00357 V=7.0 PL=0
MOVL C00358 V=7.0 PL=0
MOVL C00359 V=7.0 PL=0
MOVL C00360 V=7.0 PL=0
MOVL C00361 V=7.0 PL=0
MOVL C00362 V=7.0 PL=0
MOVL C00363 V=7.0 PL=0
MOVL C00364 V=7.0 PL=0
MOVL C00365 V=7.0 PL=0
MOVC C00366 V=7.0 ACC=20 DEC=20
MOVC C00367 V=7.0 ACC=20 DEC=20
MOVC C00368 V=7.0 ACC=20 DEC=20
MOVL C00369 V=7.0 PL=0
MOVL C00370 V=7.0 PL=0
MOVL C00371 V=7.0 PL=0
MOVL C00372 V=7.0 PL=0
MOVL C00373 V=7.0 PL=0
MOVL C00374 V=7.0 PL=0
MOVL C00375 V=7.0 PL=0
MOVL C00376 V=7.0 PL=0
MOVL C00377 V=7.0 PL=0
MOVL C00378 V=7.0 PL=0
MOVL C00379 V=7.0 PL=0
MOVL C00380 V=7.0 PL=0
MOVL C00381 V=7.0 PL=0
MOVL C00382 V=7.0 PL=0
MOVL C00383 V=7.0 PL=0
MOVL C00384 V=7.0 PL=0
MOVL C00385 V=7.0 PL=0
MOVL C00386 V=7.0 PL=0
MOVL C00387 V=7.0 PL=0
MOVL C00388 V=7.0 PL=0
ARCOF
TIMER T=30.00
*LAG10
MOVL C00389 V=11.0 PL=0
MACRO1 MJ#(0) ARGF2
ARCON
MOVL C00390 V=7.0 PL=0
MOVL C00391 V=7.0 PL=0
MOVL C00392 V=7.0 PL=0
MOVL C00393 V=7.0 PL=0
MOVL C00394 V=7.0 PL=0
MOVL C00395 V=7.0 PL=0
MOVL C00396 V=7.0 PL=0
MOVL C00397 V=7.0 PL=0
MOVL C00398 V=7.0 PL=0
MOVL C00399 V=7.0 PL=0
MOVL C00400 V=7.0 PL=0
MOVL C00401 V=7.0 PL=0
MOVL C00402 V=7.0 PL=0
MOVL C00403 V=7.0 PL=0
MOVL C00404 V=7.0 PL=0
MOVL C00405 V=7.0 PL=0
MOVL C00406 V=7.0 PL=0
MOVL C00407 V=7.0 PL=0
MOVL C00408 V=7.0 PL=0
MOVC C00409 V=7.0 ACC=20 DEC=20
MOVC C00410 V=7.0 ACC=20 DEC=20
MOVC C00411 V=7.0 ACC=20 DEC=20
MOVL C00412 V=7.0 PL=0
MOVL C00413 V=7.0 PL=0
MOVL C00414 V=7.0 PL=0
MOVL C00415 V=7.0 PL=0
MOVL C00416 V=7.0 PL=0
MOVL C00417 V=7.0 PL=0
MOVL C00418 V=7.0 PL=0
MOVL C00419 V=7.0 PL=0
MOVL C00420 V=7.0 PL=0
MOVL C00421 V=7.0 PL=0
MOVL C00422 V=7.0 PL=0
MOVL C00423 V=7.0 PL=0
MOVL C00424 V=7.0 PL=0
MOVL C00425 V=7.0 PL=0
MOVL C00426 V=7.0 PL=0
MOVL C00427 V=7.0 PL=0
MOVL C00428 V=7.0 PL=0
MOVL C00429 V=7.0 PL=0
MOVL C00430 V=7.0 PL=0
MOVL C00431 V=7.0 PL=0
ARCOF
TIMER T=30.00
*LAG11
MOVL C00432 V=11.0 PL=0
MACRO1 MJ#(0) ARGF2
ARCON
MOVL C00433 V=7.0 PL=0
MOVL C00434 V=7.0 PL=0
MOVL C00435 V=7.0 PL=0
MOVL C00436 V=7.0 PL=0
MOVL C00437 V=7.0 PL=0
MOVL C00438 V=7.0 PL=0
MOVL C00439 V=7.0 PL=0
MOVL C00440 V=7.0 PL=0
MOVL C00441 V=7.0 PL=0
MOVL C00442 V=7.0 PL=0
MOVL C00443 V=7.0 PL=0
MOVL C00444 V=7.0 PL=0
MOVL C00445 V=7.0 PL=0
MOVL C00446 V=7.0 PL=0
MOVL C00447 V=7.0 PL=0
MOVL C00448 V=7.0 PL=0
MOVL C00449 V=7.0 PL=0
MOVL C00450 V=7.0 PL=0
MOVL C00451 V=7.0 PL=0
MOVC C00452 V=7.0 ACC=20 DEC=20
MOVC C00453 V=7.0 ACC=20 DEC=20
MOVC C00454 V=7.0 ACC=20 DEC=20
MOVL C00455 V=7.0 PL=0
MOVL C00456 V=7.0 PL=0
MOVL C00457 V=7.0 PL=0
MOVL C00458 V=7.0 PL=0
MOVL C00459 V=7.0 PL=0
MOVL C00460 V=7.0 PL=0
MOVL C00461 V=7.0 PL=0
MOVL C00462 V=7.0 PL=0
MOVL C00463 V=7.0 PL=0
MOVL C00464 V=7.0 PL=0
MOVL C00465 V=7.0 PL=0
MOVL C00466 V=7.0 PL=0
MOVL C00467 V=7.0 PL=0
MOVL C00468 V=7.0 PL=0
MOVL C00469 V=7.0 PL=0
MOVL C00470 V=7.0 PL=0
MOVL C00471 V=7.0 PL=0
MOVL C00472 V=7.0 PL=0
MOVL C00473 V=7.0 PL=0
MOVL C00474 V=7.0 PL=0
ARCOF
TIMER T=30.00
*LAG12
MOVL C00475 V=11.0 PL=0
MACRO1 MJ#(0) ARGF2
ARCON
MOVL C00476 V=7.0 PL=0
MOVL C00477 V=7.0 PL=0
MOVL C00478 V=7.0 PL=0
MOVL C00479 V=7.0 PL=0
MOVL C00480 V=7.0 PL=0
MOVL C00481 V=7.0 PL=0
MOVL C00482 V=7.0 PL=0
MOVL C00483 V=7.0 PL=0
MOVL C00484 V=7.0 PL=0
MOVL C00485 V=7.0 PL=0
MOVL C00486 V=7.0 PL=0
MOVL C00487 V=7.0 PL=0
MOVL C00488 V=7.0 PL=0
MOVL C00489 V=7.0 PL=0
MOVL C00490 V=7.0 PL=0
MOVL C00491 V=7.0 PL=0
MOVL C00492 V=7.0 PL=0
MOVL C00493 V=7.0 PL=0
MOVL C00494 V=7.0 PL=0
MOVC C00495 V=7.0 ACC=20 DEC=20
MOVC C00496 V=7.0 ACC=20 DEC=20
MOVC C00497 V=7.0 ACC=20 DEC=20
MOVL C00498 V=7.0 PL=0
MOVL C00499 V=7.0 PL=0
MOVL C00500 V=7.0 PL=0
MOVL C00501 V=7.0 PL=0
MOVL C00502 V=7.0 PL=0
MOVL C00503 V=7.0 PL=0
MOVL C00504 V=7.0 PL=0
MOVL C00505 V=7.0 PL=0
MOVL C00506 V=7.0 PL=0
MOVL C00507 V=7.0 PL=0
MOVL C00508 V=7.0 PL=0
MOVL C00509 V=7.0 PL=0
MOVL C00510 V=7.0 PL=0
MOVL C00511 V=7.0 PL=0
MOVL C00512 V=7.0 PL=0
MOVL C00513 V=7.0 PL=0
MOVL C00514 V=7.0 PL=0
MOVL C00515 V=7.0 PL=0
MOVL C00516 V=7.0 PL=0
MOVL C00517 V=7.0 PL=0
ARCOF
TIMER T=30.00
*LAG13
MOVL C00518 V=11.0 PL=0
MACRO1 MJ#(0) ARGF2
ARCON
MOVL C00519 V=7.0 PL=0
MOVL C00520 V=7.0 PL=0
MOVL C00521 V=7.0 PL=0
MOVL C00522 V=7.0 PL=0
MOVL C00523 V=7.0 PL=0
MOVL C00524 V=7.0 PL=0
MOVL C00525 V=7.0 PL=0
MOVL C00526 V=7.0 PL=0
MOVL C00527 V=7.0 PL=0
MOVL C00528 V=7.0 PL=0
MOVL C00529 V=7.0 PL=0
MOVL C00530 V=7.0 PL=0
MOVL C00531 V=7.0 PL=0
MOVL C00532 V=7.0 PL=0
MOVL C00533 V=7.0 PL=0
MOVL C00534 V=7.0 PL=0
MOVL C00535 V=7.0 PL=0
MOVL C00536 V=7.0 PL=0
MOVL C00537 V=7.0 PL=0
MOVC C00538 V=7.0 ACC=20 DEC=20
MOVC C00539 V=7.0 ACC=20 DEC=20
MOVC C00540 V=7.0 ACC=20 DEC=20
MOVL C00541 V=7.0 PL=0
MOVL C00542 V=7.0 PL=0
MOVL C00543 V=7.0 PL=0
MOVL C00544 V=7.0 PL=0
MOVL C00545 V=7.0 PL=0
MOVL C00546 V=7.0 PL=0
MOVL C00547 V=7.0 PL=0
MOVL C00548 V=7.0 PL=0
MOVL C00549 V=7.0 PL=0
MOVL C00550 V=7.0 PL=0
MOVL C00551 V=7.0 PL=0
MOVL C00552 V=7.0 PL=0
MOVL C00553 V=7.0 PL=0
MOVL C00554 V=7.0 PL=0
MOVL C00555 V=7.0 PL=0
MOVL C00556 V=7.0 PL=0
MOVL C00557 V=7.0 PL=0
MOVL C00558 V=7.0 PL=0
MOVL C00559 V=7.0 PL=0
MOVL C00560 V=7.0 PL=0
ARCOF
TIMER T=30.00
*LAG14
MOVL C00561 V=11.0 PL=0
MACRO1 MJ#(0) ARGF2
ARCON
MOVL C00562 V=7.0 PL=0
MOVL C00563 V=7.0 PL=0
MOVL C00564 V=7.0 PL=0
MOVL C00565 V=7.0 PL=0
MOVL C00566 V=7.0 PL=0
MOVL C00567 V=7.0 PL=0
MOVL C00568 V=7.0 PL=0
MOVL C00569 V=7.0 PL=0
MOVL C00570 V=7.0 PL=0
MOVL C00571 V=7.0 PL=0
MOVL C00572 V=7.0 PL=0
MOVL C00573 V=7.0 PL=0
MOVL C00574 V=7.0 PL=0
MOVL C00575 V=7.0 PL=0
MOVL C00576 V=7.0 PL=0
MOVL C00577 V=7.0 PL=0
MOVL C00578 V=7.0 PL=0
MOVL C00579 V=7.0 PL=0
MOVL C00580 V=7.0 PL=0
MOVC C00581 V=7.0 ACC=20 DEC=20
MOVC C00582 V=7.0 ACC=20 DEC=20
MOVC C00583 V=7.0 ACC=20 DEC=20
MOVL C00584 V=7.0 PL=0
MOVL C00585 V=7.0 PL=0
MOVL C00586 V=7.0 PL=0
MOVL C00587 V=7.0 PL=0
MOVL C00588 V=7.0 PL=0
MOVL C00589 V=7.0 PL=0
MOVL C00590 V=7.0 PL=0
MOVL C00591 V=7.0 PL=0
MOVL C00592 V=7.0 PL=0
MOVL C00593 V=7.0 PL=0
MOVL C00594 V=7.0 PL=0
MOVL C00595 V=7.0 PL=0
MOVL C00596 V=7.0 PL=0
MOVL C00597 V=7.0 PL=0
MOVL C00598 V=7.0 PL=0
MOVL C00599 V=7.0 PL=0
MOVL C00600 V=7.0 PL=0
MOVL C00601 V=7.0 PL=0
MOVL C00602 V=7.0 PL=0
MOVL C00603 V=7.0 PL=0
ARCOF
TIMER T=30.00
*LAG15
MOVL C00604 V=11.0 PL=0
MACRO1 MJ#(0) ARGF2
ARCON
MOVL C00605 V=7.0 PL=0
MOVL C00606 V=7.0 PL=0
MOVL C00607 V=7.0 PL=0
MOVL C00608 V=7.0 PL=0
MOVL C00609 V=7.0 PL=0
MOVL C00610 V=7.0 PL=0
MOVL C00611 V=7.0 PL=0
MOVL C00612 V=7.0 PL=0
MOVL C00613 V=7.0 PL=0
MOVL C00614 V=7.0 PL=0
MOVL C00615 V=7.0 PL=0
MOVL C00616 V=7.0 PL=0
MOVL C00617 V=7.0 PL=0
MOVL C00618 V=7.0 PL=0
MOVL C00619 V=7.0 PL=0
MOVL C00620 V=7.0 PL=0
MOVL C00621 V=7.0 PL=0
MOVL C00622 V=7.0 PL=0
MOVL C00623 V=7.0 PL=0
MOVC C00624 V=7.0 ACC=20 DEC=20
MOVC C00625 V=7.0 ACC=20 DEC=20
MOVC C00626 V=7.0 ACC=20 DEC=20
MOVL C00627 V=7.0 PL=0
MOVL C00628 V=7.0 PL=0
MOVL C00629 V=7.0 PL=0
MOVL C00630 V=7.0 PL=0
MOVL C00631 V=7.0 PL=0
MOVL C00632 V=7.0 PL=0
MOVL C00633 V=7.0 PL=0
MOVL C00634 V=7.0 PL=0
MOVL C00635 V=7.0 PL=0
MOVL C00636 V=7.0 PL=0
MOVL C00637 V=7.0 PL=0
MOVL C00638 V=7.0 PL=0
MOVL C00639 V=7.0 PL=0
MOVL C00640 V=7.0 PL=0
MOVL C00641 V=7.0 PL=0
MOVL C00642 V=7.0 PL=0
MOVL C00643 V=7.0 PL=0
MOVL C00644 V=7.0 PL=0
MOVL C00645 V=7.0 PL=0
MOVL C00646 V=7.0 PL=0
ARCOF
TIMER T=30.00
MOVL C00647 V=11.0 PL=0
MOVJ C00648 VJ=0.78
END
